Fanuc KAREL source: KT00314.KL

PROGRAM KT00314
%NOLOCKGROUP
VAR
  P1: POSITION
  P2: JOINTPOS
  OUT: BOOLEAN
BEGIN
  OUT = P1 <> P2
END KT00314
